(* IEC 61131-3 sources: tsplc/packages/build/tests/fixtures/raw-st/src/filling/FB_FillingStation, 2 files *)

(* ---- declaration.st ---- *)
FUNCTION_BLOCK FB_FillingStation
VAR
	State : E_StationState := E_StationState.Idle;
	Completed : UDINT;
END_VAR

(* ---- FB_FillingStation.implementation.st ---- *)
CASE State OF
	E_StationState.Idle: State := E_StationState.Working;
	E_StationState.Working:
		Completed := Completed + 1;
		State := E_StationState.Idle;
END_CASE
